// TIA Portal V21 export
// export: Created 2026-08-21T20:18:55.7123431Z, ExportSetting None, DisplayName Totally Integrated Automation Portal, DisplayVersion V21, DisplayName STEP 7 Professional, DisplayVersion V21, DisplayName STEP 7 Safety, DisplayVersion V21, DisplayName Tech WebApplication, DisplayVersion V21, DisplayName WinCC Basic/Comfort/Advanced, DisplayVersion V21, DisplayName WinCC Professional, DisplayVersion V21, DisplayName WinCC Unified, DisplayVersion V21
TYPE "ScaVal_Raw"
   STRUCT
      High : DInt := 32767;   // High Value
      Low : DInt := -32768;   // Low Value
   END_STRUCT;
END_TYPE
